{attribute 'OPC.UA.DA.StructuredType' := '1'}
TYPE ST_HeatPumpBufferState :
STRUCT
	fMidTemperature 	: REAL;
END_STRUCT
END_TYPE

(* stored: Version 1.1.0.1
   DUT ST_HeatPumpBufferState: Id {f07d6861-270a-4dbd-875a-4a83b5c7c554} *)
